FUNCTION_BLOCK F (* Positive: exit guards read a variable that this scan's algorithm has just assigned, which is not dispatch *)
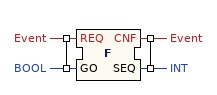
  EVENT_INPUT
    REQ WITH GO;
  END_EVENT
  EVENT_OUTPUT
    CNF WITH SEQ;
  END_EVENT
  VAR_INPUT
    GO : BOOL;
  END_VAR
  VAR_OUTPUT
    SEQ : INT;
  END_VAR
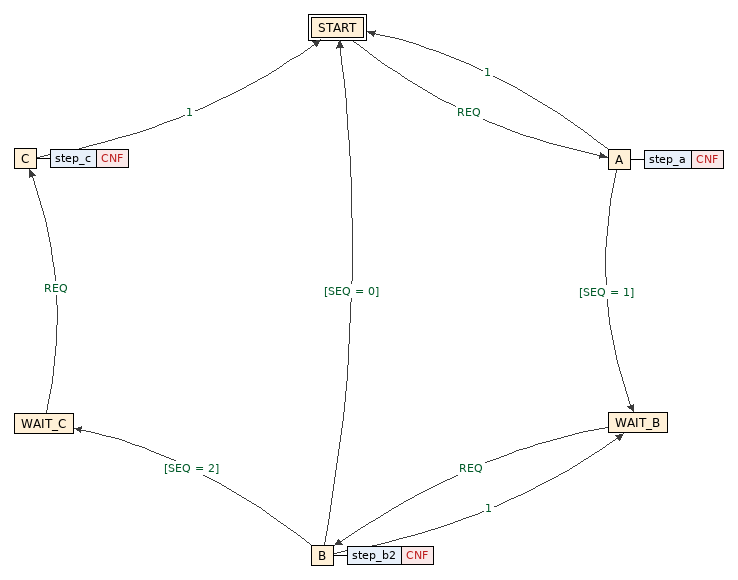
  EC_STATES
    START;
    A : step_a -> CNF;
    WAIT_B;
    B : step_b2 -> CNF;
    WAIT_C;
    C : step_c -> CNF;
  END_STATES
  EC_TRANSITIONS
    START TO A := REQ;
    A TO WAIT_B := [SEQ = 1];
    A TO START := 1;
    WAIT_B TO B := REQ;
    B TO WAIT_C := [SEQ = 2];
    B TO START := [SEQ = 0];
    B TO WAIT_B := 1;
    WAIT_C TO C := REQ;
    C TO START := 1;
  END_TRANSITIONS
  ALGORITHM step_a IN ST:
SEQ := 0;
IF GO THEN
  SEQ := 1;
END_IF;
  END_ALGORITHM
  ALGORITHM step_b2 IN ST:
IF GO THEN
  SEQ := 2;
ELSE
  SEQ := 0;
END_IF;
  END_ALGORITHM
  ALGORITHM step_c IN ST:
SEQ := 0;
  END_ALGORITHM
END_FUNCTION_BLOCK
